Yaskawa INFORM job: 123.JBI

/JOB
//NAME 123
//POS
///NPOS 42,42,42,0,0,0
///TOOL 0
///POSTYPE PULSE
///PULSE
C00000=-286,-101165,-84213,3710,-80189,-1933
C00001=-285,-101145,-84203,3591,-80198,-1944
C00002=-285,-101145,-84203,3591,-80198,-1944
C00003=-89705,50615,23938,-6742,-70649,29246
C00004=-104514,76177,-5240,-73154,-45601,55743
C00005=-105404,73854,-8195,-73415,-45851,56215
C00006=-103220,74581,-7274,-74028,-44814,55869
C00007=-103220,73831,-7282,-73660,-44930,55635
C00008=-103220,73831,-7282,-73660,-44930,55635
C00009=-103220,73831,-7282,-73660,-44930,55635
C00010=-103304,76029,-4494,-73068,-45156,55285
C00011=-103413,77324,-4138,-73456,-45070,55570
C00012=-102803,71565,-11546,-75244,-44287,56503
C00013=-102803,65225,-11333,-71963,-45337,54415
C00014=-104478,64301,-12450,-71622,-46129,54741
C00015=-101589,61882,-22935,-77812,-43156,57692
C00016=-101774,63036,-21526,-77448,-43313,57529
C00017=-102511,62694,-22140,-77345,-43621,57720
C00018=-102396,66494,-17467,-76424,-43803,57118
C00019=-102396,59611,-17179,-72748,-44895,54798
C00020=-104285,64730,-19843,-76208,-44578,57634
C00021=-104859,63785,-20571,-75932,-44871,57662
C00022=-104538,60478,-24614,-76840,-44509,58126
C00023=-103872,60156,-25004,-77200,-44170,58118
C00024=-104477,59871,-25349,-77005,-44444,58210
C00025=-103333,60361,-24457,-77196,-43968,57927
C00026=-102823,61345,-23264,-77178,-43780,57739
C00027=-102591,62916,-21584,-77045,-43725,57579
C00028=-102591,59617,-21542,-75304,-44186,56488
C00029=-103891,49710,-33174,-76848,-44266,57908
C00030=-103673,54286,-32569,-78960,-43688,59154
C00031=-103647,52324,-34326,-79047,-43660,59199
C00032=-103475,50803,-36106,-79453,-43512,59390
C00033=-102931,50687,-36238,-79732,-43253,59369
C00034=-102427,52656,-33930,-79539,-43103,59068
C00035=-102331,53867,-32504,-79311,-43112,58894
C00036=-102094,51906,-34812,-79859,-42914,59148
C00037=-101420,51023,-35597,-80208,-42595,59124
C00038=-101178,53725,-32870,-80009,-42539,58918
C00039=-60698,-7215,-10633,-28437,-86038,24832
C00040=-285,-101145,-84203,3591,-80198,-1944
C00041=-285,-101145,-84203,3591,-80198,-1944
BC00000=570125
BC00001=570127
BC00002=847209
BC00003=847209
BC00004=847208
BC00005=847208
BC00006=847208
BC00007=847208
BC00008=847208
BC00009=847208
BC00010=847208
BC00011=847208
BC00012=847208
BC00013=847208
BC00014=847208
BC00015=847208
BC00016=847208
BC00017=847208
BC00018=847207
BC00019=847207
BC00020=847207
BC00021=847207
BC00022=847207
BC00023=847207
BC00024=847207
BC00025=847207
BC00026=847207
BC00027=847207
BC00028=847207
BC00029=847207
BC00030=847207
BC00031=847207
BC00032=847207
BC00033=847207
BC00034=847207
BC00035=847207
BC00036=847207
BC00037=847207
BC00038=847207
BC00039=847208
BC00040=847209
BC00041=570127
EC00000=1,4
EC00001=3,-5
EC00002=3,-5
EC00003=3,-5
EC00004=3,-5
EC00005=3,-5
EC00006=3,-5
EC00007=3,-5
EC00008=3,-5
EC00009=3,-5
EC00010=3,-5
EC00011=3,-5
EC00012=3,-5
EC00013=3,-5
EC00014=3,-5
EC00015=3,-5
EC00016=3,-5
EC00017=3,-5
EC00018=3,-5
EC00019=3,-5
EC00020=3,-5
EC00021=3,-5
EC00022=3,-5
EC00023=3,-5
EC00024=3,-5
EC00025=3,-5
EC00026=3,-5
EC00027=3,-5
EC00028=3,-5
EC00029=3,-5
EC00030=3,-5
EC00031=3,-5
EC00032=3,-5
EC00033=3,-5
EC00034=3,-5
EC00035=3,-5
EC00036=3,-5
EC00037=3,-5
EC00038=3,-5
EC00039=3,-5
EC00040=3,-5
EC00041=3,-5
//INST
///DATE 2025/01/10 11:19
///ATTR SC,RW
///GROUP1 RB1,BS1
///GROUP2 ST3
NOP
MOVJ C00000 BC00000 VJ=0.78 DEC=20  +MOVJ EC00000 VJ=0.78
MOVJ C00001 BC00001 VJ=0.78  +MOVJ EC00001 VJ=0.78
MOVJ C00002 BC00002 VJ=90.00  +MOVJ EC00002 VJ=0.78
MOVJ C00003 BC00003 VJ=90.00  +MOVJ EC00003 VJ=0.78
MOVJ C00004 BC00004 VJ=90.00  +MOVJ EC00004 VJ=0.78
MACRO1 MJ#(0) ARGF1
MOVL C00005 BC00005 V=2.5  +MOVJ EC00005 VJ=0.78
MOVL C00006 BC00006 V=3.3  +MOVJ EC00006 VJ=0.78
MOVJ C00007 BC00007 VJ=20.00  +MOVJ EC00007 VJ=20.00
MOVJ C00008 BC00008 VJ=20.00  +MOVJ EC00008 VJ=20.00
MOVJ C00009 BC00009 VJ=20.00  +MOVJ EC00009 VJ=20.00
MOVJ C00010 BC00010 VJ=20.00  +MOVJ EC00010 VJ=20.00
MOVJ C00011 BC00011 VJ=20.00  +MOVJ EC00011 VJ=20.00
MOVL C00012 BC00012 V=5.0  +MOVJ EC00012 VJ=20.00
MOVJ C00013 BC00013 VJ=20.00  +MOVJ EC00013 VJ=20.00
MOVJ C00014 BC00014 VJ=20.00  +MOVJ EC00014 VJ=20.00
MOVJ C00015 BC00015 VJ=20.00  +MOVJ EC00015 VJ=20.00
MOVL C00016 BC00016 V=5.0  +MOVJ EC00016 VJ=20.00
MOVL C00017 BC00017 V=3.3  +MOVJ EC00017 VJ=20.00
MOVL C00018 BC00018 V=3.3  +MOVJ EC00018 VJ=20.00
MOVJ C00019 BC00019 VJ=90.00  +MOVJ EC00019 VJ=20.00
MOVJ C00020 BC00020 VJ=90.00  +MOVJ EC00020 VJ=90.00
MOVL C00021 BC00021 V=3.3  +MOVJ EC00021 VJ=90.00
MOVL C00022 BC00022 V=5.0  +MOVJ EC00022 VJ=90.00
MOVC C00023 BC00023 V=3.3  +MOVJ EC00023 VJ=90.00
MOVC C00024 BC00024 V=3.3  +MOVJ EC00024 VJ=90.00
MOVC C00025 BC00025 V=3.3  +MOVJ EC00025 VJ=90.00
MOVC C00026 BC00026 V=3.3  +MOVJ EC00026 VJ=90.00
MOVC C00027 BC00027 V=3.3  +MOVJ EC00027 VJ=90.00
MOVJ C00028 BC00028 VJ=90.00  +MOVJ EC00028 VJ=90.00
MOVJ C00029 BC00029 VJ=90.00  +MOVJ EC00029 VJ=90.00
MOVJ C00030 BC00030 VJ=90.00  +MOVJ EC00030 VJ=90.00
MOVL C00031 BC00031 V=3.3  +MOVJ EC00031 VJ=90.00
MOVL C00032 BC00032 V=3.3  +MOVJ EC00032 VJ=90.00
MOVC C00033 BC00033 V=3.3  +MOVJ EC00033 VJ=90.00
MOVC C00034 BC00034 V=3.3  +MOVJ EC00034 VJ=90.00
MOVC C00035 BC00035 V=3.3  +MOVJ EC00035 VJ=90.00
MOVC C00036 BC00036 V=3.3  +MOVJ EC00036 VJ=90.00
MOVC C00037 BC00037 V=3.3  +MOVJ EC00037 VJ=90.00
MOVC C00038 BC00038 V=3.3  +MOVJ EC00038 VJ=90.00
MOVJ C00039 BC00039 VJ=90.00  +MOVJ EC00039 VJ=90.00
MOVJ C00040 BC00040 VJ=90.00  +MOVJ EC00040 VJ=90.00
MOVJ C00041 BC00041 VJ=90.00  +MOVJ EC00041 VJ=90.00
END
